(* PLC project probe.project, CODESYS CODESYS V3.5 SP17 Patch 3 *)
(* stored: creationDateTime 2026-10-20T03:54:26.7835114, modificationDateTime 1601-01-01T03:00:00 *)

FUNCTION_BLOCK FB_ProbeLd
  VAR_INPUT
    xStart : BOOL;
    xStop : BOOL;
    xPermit : BOOL;
    iSp : INT;
  END_VAR
  VAR_OUTPUT
    xRun : BOOL;
    iOut : INT;
    xMoved : BOOL;
    xRunInv : BOOL;
  END_VAR
  VAR  (* added by the conversion: wires and edge detectors of the diagram *)
    R_TRIG1 : R_TRIG;
    F_TRIG2 : F_TRIG;
  END_VAR

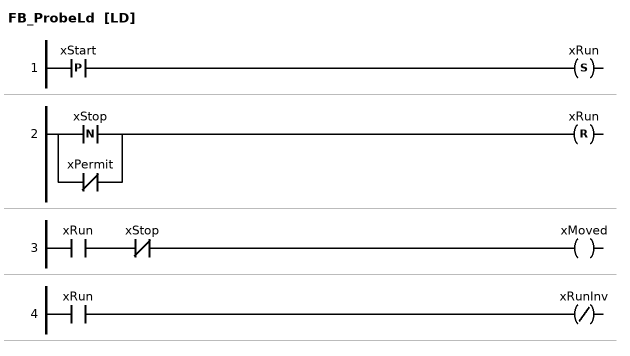
(* LD diagram, written out as Structured Text *)
(* --- network: Пуск по фронту --- *)
R_TRIG1(CLK := xStart);
IF R_TRIG1.Q THEN xRun := TRUE; END_IF;
(* --- network: Стоп по спаду или без разрешения --- *)
F_TRIG2(CLK := xStop);
IF F_TRIG2.Q OR NOT xPermit THEN xRun := FALSE; END_IF;
(* --- network: Последовательная цепь --- *)
xMoved := xRun AND NOT xStop;
(* --- network: Инверсная катушка --- *)
xRunInv := NOT xRun;
END_FUNCTION_BLOCK
